// TIA Portal V21 export
// export: Created 2026-11-21T23:19:38.16006Z, ExportSetting WithDefaults, DisplayName Totally Integrated Automation Portal, DisplayVersion V21 Update 3, DisplayName STEP 7 Professional, DisplayVersion V21 Update 3, DisplayName STEP 7 Safety, DisplayVersion V21, DisplayName Tech WebApplication, DisplayVersion V21, DisplayName WinCC Basic/Comfort/Advanced, DisplayVersion V21 Update 3, DisplayName WinCC Unified, DisplayVersion V21 Update 3
Cycle "Default cycle 1"  CycleTime=2, CycleUnit=Second, StartingPoint=****-**-**T**:**:**
